Staubli VAL3: setMark.pgx

public program setMark(string x_sKey, num x_nIndex)
begin

  trajTemp:tTrajItem[x_sKey].pPointItem[x_nIndex].bMarked=!trajTemp:tTrajItem[x_sKey].pPointItem[x_nIndex].bMarked
//  if trajTemp:tTrajItem[x_sKey].pPointItem[x_nIndex].bMarked
//    savedata:nMarkIndex[x_nIndex]=1
//  else
//    savedata:nMarkIndex[x_nIndex]=-1
//  endIf

end
